// TIA Portal V19 export
VAR_GLOBAL   // PLC tag table "R2_OUT"
   "ByteOUT :0 R2" AT %QB206 : Byte;   // System Bits 1
   "ByteOUT :1 R2" AT %QB207 : Byte;   // System Bits 2
   "ByteOUT :2 R2" AT %QB208 : Byte;   // Signals
   "ByteOUT :3 R2" AT %QB209 : Byte;   // Signals
   "ByteOUT :4 R2" AT %QB210 : Byte;   // CMD
   "ByteOUT :5 R2" AT %QB211 : Byte;   // CMD
   "ByteOUT :6 R2" AT %QB212 : Byte;   // X
   "ByteOUT :7 R2" AT %QB213 : Byte;   // X
   "ByteOUT :8 R2" AT %QB214 : Byte;   // Y
   "ByteOUT :9 R2" AT %QB215 : Byte;   // Y
   "ByteOUT :10 R2" AT %QB216 : Byte;   // Z
   "ByteOUT :11 R2" AT %QB217 : Byte;   // Z
   "ByteOUT :12 R2" AT %QB218 : Byte;
   "ByteOUT :13 R2" AT %QB219 : Byte;
   "ByteOUT :14 R2" AT %QB220 : Byte;
   "ByteOUT :15 R2" AT %QB221 : Byte;
   "ByteOUT :16 R2" AT %QB222 : Byte;
   "ByteOUT :17 R2" AT %QB223 : Byte;
   "ByteOUT :18 R2" AT %QB224 : Byte;
   "ByteOUT :19 R2" AT %QB225 : Byte;
   "ByteOUT :20 R2" AT %QB226 : Byte;
   "ByteOUT :21 R2" AT %QB227 : Byte;
   "ByteOUT :22 R2" AT %QB228 : Byte;
   "ByteOUT :23 R2" AT %QB229 : Byte;
   "ByteOUT :24 R2" AT %QB230 : Byte;
   "ByteOUT :25 R2" AT %QB231 : Byte;
   "ByteOUT :26 R2" AT %QB232 : Byte;
   "ByteOUT :27 R2" AT %QB233 : Byte;
   "ByteOUT :28 R2" AT %QB234 : Byte;
   "ByteOUT :29 R2" AT %QB235 : Byte;
   "ByteOUT :30 R2" AT %QB236 : Byte;
   "ByteOUT :31 R2" AT %QB237 : Byte;
   "ByteOUT :32 R2" AT %QB238 : Byte;
   "ByteOUT :33 R2" AT %QB239 : Byte;
   "ByteOUT :34 R2" AT %QB240 : Byte;
   "ByteOUT :35 R2" AT %QB241 : Byte;
   "ByteOUT :36 R2" AT %QB242 : Byte;
   "ByteOUT :37 R2" AT %QB243 : Byte;
   "ByteOUT :38 R2" AT %QB244 : Byte;
   "ByteOUT :39 R2" AT %QB245 : Byte;
   "ByteOUT :40 R2" AT %QB246 : Byte;
   "ByteOUT :41 R2" AT %QB247 : Byte;
   "ByteOUT :42 R2" AT %QB248 : Byte;
   "ByteOUT :43 R2" AT %QB249 : Byte;
   "ByteOUT :44 R2" AT %QB250 : Byte;
   "ByteOUT :45 R2" AT %QB251 : Byte;
   "ByteOUT :46 R2" AT %QB252 : Byte;
   "ByteOUT :47 R2" AT %QB253 : Byte;
   "ByteOUT :48 R2" AT %QB254 : Byte;
   "ByteOUT :49 R2" AT %QB255 : Byte;
   "ByteOUT :50 R2" AT %QB256 : Byte;
   "ByteOUT :51 R2" AT %QB257 : Byte;
   "ByteOUT :52 R2" AT %QB258 : Byte;
   "ByteOUT :53 R2" AT %QB259 : Byte;
   "ByteOUT :54 R2" AT %QB260 : Byte;
   "ByteOUT :55 R2" AT %QB261 : Byte;
   "ByteOUT :56 R2" AT %QB262 : Byte;
   "ByteOUT :57 R2" AT %QB263 : Byte;
   "ByteOUT :58 R2" AT %QB264 : Byte;
   "ByteOUT :59 R2" AT %QB265 : Byte;
   "ByteOUT :60 R2" AT %QB266 : Byte;
   "ByteOUT :61 R2" AT %QB267 : Byte;
   "ByteOUT :62 R2" AT %QB268 : Byte;
   "ByteOUT :63 R2" AT %QB269 : Byte;
END_VAR
